SUBAPPLICATION logiBUS_AI_MVA_Scaled_OPC (* Analog-Eingang in mV (Pin), feste Umrechnung OUT = mV * SCALE + OFFSET, Publish mV und Wert (ohne VT) *)
  (* Standard: 61499-2; Description: Copyright (c) 2026 Meisterschulen am Ostbahnhof This program and the accompanying materials are made available under the terms of the Eclipse Public License 2.0 which is available at https://www.eclipse.org/legal/epl-2.0/ SPDX-License-Identifier: EPL-2.0 *)
  (* Version 1.0, 2026-11-15, Franz Höpfinger, Meisterschulen am Ostbahnhof, initial API and implementation and/or initial documentation *)
  PACKAGE MyLib::sys;
  IMPORT logiBUS::io::AI::logiBUS_AI;
  IMPORT logiBUS::io::AI::logiBUS_AI_S;
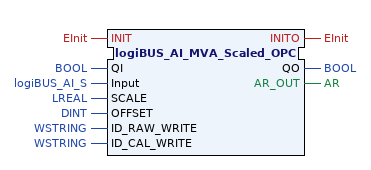
  EVENT_INPUT
    INIT : EInit; (* Initialization Request *)
  END_EVENT
  EVENT_OUTPUT
    INITO : EInit; (* Initialization Confirm *)
  END_EVENT
  VAR_INPUT
    QI : BOOL := TRUE; (* Quality Input - TRUE to enable service *)
    Input : logiBUS::io::AI::logiBUS_AI_S := logiBUS_AI::Invalid; (* Identify the Input AnalogInput_I1..I8 *)
    SCALE : LREAL := LREAL#1.0; (* Faktor je mV am Pin *)
    OFFSET : DINT := DINT#0; (* Offset nach dem Faktor *)
    ID_RAW_WRITE : WSTRING; (* Pin-mV (REAL, ACTION=PUBLISH) *)
    ID_CAL_WRITE : WSTRING; (* Umgerechneter Wert (REAL, ACTION=PUBLISH) *)
  END_VAR
  VAR_OUTPUT
    QO : BOOL; (* Quality Output - TRUE if service executed successfully *)
  END_VAR
  PLUGS
    AR_OUT : adapter::types::unidirectional::AR; (* Umgerechneter Wert *)
  END_PLUGS
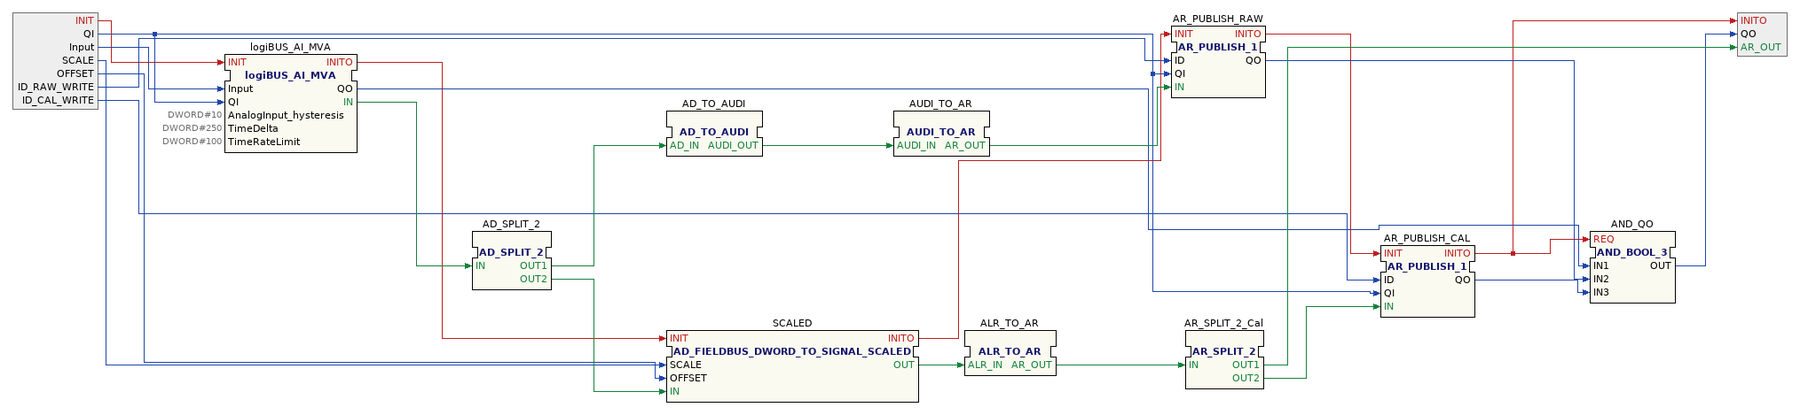
  FBS
    logiBUS_AI_MVA : logiBUS::io::AI::logiBUS_AI_MVA(AnalogInput_hysteresis := DWORD#10, TimeDelta := DWORD#250, TimeRateLimit := DWORD#100);
    AD_SPLIT_2 : adapter::events::unidirectional::AD_SPLIT_2;
    AD_TO_AUDI : adapter::conversion::unidirectional::AD_TO_AUDI;
    AUDI_TO_AR : adapter::conversion::unidirectional::AUDI_TO_AR;
    AR_PUBLISH_RAW : adapter::net::AR_PUBLISH_1;
    SCALED : logiBUS::signalprocessing::fieldbus::AD_FIELDBUS_DWORD_TO_SIGNAL_SCALED;
    ALR_TO_AR : adapter::conversion::unidirectional::ALR_TO_AR;
    AR_SPLIT_2_Cal : adapter::events::unidirectional::AR_SPLIT_2;
    AR_PUBLISH_CAL : adapter::net::AR_PUBLISH_1;
    AND_QO : iec61131::booleanOperators::AND_BOOL_3;
  END_FBS
  EVENT_CONNECTIONS
    INIT TO logiBUS_AI_MVA.INIT;
    logiBUS_AI_MVA.INITO TO SCALED.INIT;
    SCALED.INITO TO AR_PUBLISH_RAW.INIT;
    AR_PUBLISH_RAW.INITO TO AR_PUBLISH_CAL.INIT;
    AR_PUBLISH_CAL.INITO TO INITO;
    AR_PUBLISH_CAL.INITO TO AND_QO.REQ;
  END_CONNECTIONS
  DATA_CONNECTIONS
    Input TO logiBUS_AI_MVA.Input;
    QI TO logiBUS_AI_MVA.QI;
    SCALE TO SCALED.SCALE;
    OFFSET TO SCALED.OFFSET;
    ID_RAW_WRITE TO AR_PUBLISH_RAW.ID;
    QI TO AR_PUBLISH_RAW.QI;
    ID_CAL_WRITE TO AR_PUBLISH_CAL.ID;
    QI TO AR_PUBLISH_CAL.QI;
    logiBUS_AI_MVA.QO TO AND_QO.IN1;
    AR_PUBLISH_RAW.QO TO AND_QO.IN2;
    AR_PUBLISH_CAL.QO TO AND_QO.IN3;
    AND_QO.OUT TO QO;
  END_CONNECTIONS
  ADAPTER_CONNECTIONS
    logiBUS_AI_MVA.IN TO AD_SPLIT_2.IN;
    AD_SPLIT_2.OUT1 TO AD_TO_AUDI.AD_IN;
    AD_TO_AUDI.AUDI_OUT TO AUDI_TO_AR.AUDI_IN;
    AUDI_TO_AR.AR_OUT TO AR_PUBLISH_RAW.IN;
    AD_SPLIT_2.OUT2 TO SCALED.IN;
    SCALED.OUT TO ALR_TO_AR.ALR_IN;
    ALR_TO_AR.AR_OUT TO AR_SPLIT_2_Cal.IN;
    AR_SPLIT_2_Cal.OUT1 TO AR_OUT;
    AR_SPLIT_2_Cal.OUT2 TO AR_PUBLISH_CAL.IN;
  END_CONNECTIONS
END_SUBAPPLICATION
